(* IEC 61131-3 sources: trust-platform/editors/vscode/media/examples/raspberry-pi/src, 2 files *)

(* ---- config.st ---- *)
CONFIGURATION Config
RESOURCE MainRes ON PLC
    TASK MainTask (INTERVAL := T#10ms, PRIORITY := 1);
    PROGRAM Main WITH MainTask : Main;
END_RESOURCE
END_CONFIGURATION

(* ---- Main.st ---- *)
PROGRAM Main
VAR
    output_on : BOOL;
    ticks     : DINT;
END_VAR
    ticks := ticks + 1;
    output_on := (ticks MOD 100) < 50;
END_PROGRAM
